(*
SPDX-FileCopyrightText: © 2026 Oleksandr Tiutyk <trofimich@gmail.com>
SPDX-License-Identifier: MIT
License: https://opensource.org/license/mit
*)

(*!
<summary>Exposes diagnostics for a missing workflow variable.</summary>
<description>
Reports when a required workflow variable cannot be found in the current activity or workflow scope. Dynamic
copies are explicitly registered by Clone after construction; plain __NEW does not transfer ownership to the
task manager.
</description>
*)

{attribute 'enable_dynamic_creation'}
{attribute 'no_explicit_call' := 'do not call this function block directly'}
FUNCTION_BLOCK WorkflowVariableNotFoundException EXTENDS TOF_Core.GeneralException
	IMPLEMENTS IWorkflowVariableNotFoundException
VAR_STAT
	{attribute 'hide'} 
	_ClassName : STRING := __POUNAME();
END_VAR

(*!
<summary>Borrows the initialized class name used in diagnostics.</summary>
<description>
Returns initialized metadata storage without allocation. Callers must not modify the returned string.
Derived function blocks must use distinct initialized static storage when overriding this metadata.
</description>
*)
{attribute 'monitoring' := 'call'}
PROPERTY ClassName : REFERENCE TO STRING
GET
ClassName REF= _ClassName;
END_GET
END_PROPERTY

(*!
<summary>Creates a task-owned copy of this exception and its diagnostic payload.</summary>
<description>
Registers the newly constructed instance before copying payload, outside FB_init. Registration failure
releases the unregistered instance and raises a terminal error; copy failure leaves the registered instance
owned by the task manager for cleanup. Custom overrides must follow the same ownership sequence. The returned
reference is borrowed until task cleanup and must not be deleted by the caller.
</description>
*)
METHOD Clone : TOF_Core.IObject
VAR
	exceptionClone : POINTER TO WorkflowVariableNotFoundException;
END_VAR
exceptionClone := __NEW(WorkflowVariableNotFoundException);

IF exceptionClone = 0 THEN
	TOF_Core.DynamicMemoryManager.RaiseAllocationFailure();
END_IF

TOF_Core.DynamicMemoryManager.RegisterAutoDisposedObject(autoDisposedObject := exceptionClone^);

exceptionClone^.CopyGeneralFields(sourceException := THIS^);

Clone := exceptionClone^;
END_METHOD

(*!
<summary>Provides the library namespace used in diagnostics.</summary>
<description>Returns borrowed read-only namespace storage; do not modify the referenced string.</description>
*)
{attribute 'monitoring' := 'call'}
PROPERTY NamespaceName : REFERENCE TO STRING
GET
NamespaceName REF= CurrentNamespace.Name;
END_GET
END_PROPERTY

(*!
<summary>Reports the size of this concrete instance in bytes.</summary>
*)
{attribute 'monitoring' := 'call'}
PROPERTY SelfSize : ULINT
GET
SelfSize := XSIZEOF(THIS^);
END_GET
END_PROPERTY

(*!
<summary>Raises an exception describing the missing workflow variable.</summary>
<description>
Borrows message read-only for this call and formats diagnostic text without heap allocation during message
preparation.
</description>
<param name="sourceNamespaceName">Namespace of the caller.</param>
<param name="sourceClassName">Class name of the caller.</param>
<param name="sourcePOUName">POU name of the caller.</param>
<param name="sourcePosition">Source position of the caller.</param>
<param name="message">Diagnostic explanation.</param>
*)
METHOD Throw
VAR_INPUT
	sourceNamespaceName : STRING;
	sourceClassName : STRING;
	sourcePOUName : STRING;
	sourcePosition : STRING;
END_VAR
VAR_IN_OUT CONSTANT
	message : TOF_Core.ERROR_MESSAGE;
END_VAR
InternalThrow(
	sourceNamespaceName := sourceNamespaceName,
	sourceClassName := sourceClassName,
	sourcePOUName := sourcePOUName,
	sourcePosition := sourcePosition,
	message := message,
	errorCode := 0,
	innerException := 0
);
END_METHOD

END_FUNCTION_BLOCK

(* stored: Version 1.1.0.1
   POU WorkflowVariableNotFoundException: Id {b55861eb-5eed-49b6-afac-e9bf81d71e38}, SpecialFunc None
   Property ClassName: Id {82b7d44c-eae1-4dde-9670-6ebec99667b7}
   Get Get: Id {d3588156-bee9-49b6-9a6c-04ea18d90604}
   Method Clone: Id {4406c442-56b0-4754-b0e5-b1f015e89840}
   Property NamespaceName: Id {1c8fb75c-bfa0-4573-bb2f-b02b01e4b6d8}
   Get Get: Id {6cd1c55a-227f-47b5-b006-5d766018e063}
   Property SelfSize: Id {1fb58c0b-ff84-496a-bc07-47ad4453e478}
   Get Get: Id {e2f84cbc-8bfc-480a-a107-4c88a44861cd}
   Method Throw: Id {26879042-1e82-421e-9d95-84683b3b975c} *)
